(* IEC 61131-3 sources: plc-st-coding-agent/progress/evidence/f14_v14_remaining_20261113/jobs/custom_minimax-m27 (part 9) *)

(* ---- self-medium-04.raw_candidate_01.st ---- *)
FUNCTION_BLOCK FB
VAR_INPUT
    startBtn  : BOOL;
    resetBtn  : BOOL;
    doneSensor: BOOL;
    targetVol : REAL;
    flowVol   : REAL;
END_VAR
VAR_OUTPUT
    valveOpen : BOOL;
    fillsToday: INT;
END_VAR
VAR
    state           : INT;        // 0=IDLE, 1=FILLING, 2=PENDING
    prev_startBtn   : BOOL;
    prev_resetBtn   : BOOL;
    prev_valveOpen  : BOOL;
    pendingConfirm  : BOOL;
    accumulatedVol  : REAL;
    rising_startBtn : BOOL;
    rising_resetBtn : BOOL;
    tmp_doConfirm   : BOOL;
END_VAR

// ENGINEERING_CONTRACT
// States: IDLE(0), FILLING(1), PENDING(2)
// Outputs: valveOpen (BOOL, hold open during FILLING until target reached or reset)
//          fillsToday (INT, hold-until-confirm count, saturation at 32767)
// Confirmed fills increment fillsToday by 1 per bottle, cleared on reset
// ResetBtn rising edge (rising_resetBtn) has absolute priority; clears all state
// StartBtn rising edge (rising_startBtn) in IDLE or PENDING starts new bottle
// Confirmation checks doneSensor at valve-close scan; clears pendingConfirm after
// No hidden timers; all state in VAR; explicit edge detection via prev_* vars

(* CONTRACT_RULES [] *)

rising_startBtn := startBtn AND NOT prev_startBtn;
rising_resetBtn := resetBtn  AND NOT prev_resetBtn;

// PUB001: Reset takes priority - ignore everything else this scan
IF rising_resetBtn THEN
    pendingConfirm := FALSE;
    accumulatedVol := 0.0;
    valveOpen      := FALSE;
    fillsToday     := 0;
    prev_startBtn  := startBtn;
    prev_resetBtn  := resetBtn;
    prev_valveOpen := valveOpen;
    RETURN;
END_IF;

// PUB002: Start new bottle when startBtn rises (idle or waiting confirmation)
IF rising_startBtn AND (state = 0 OR state = 2) THEN
    state           := 1;          // FILLING
    pendingConfirm  := FALSE;      // cancel previous pending if any
    accumulatedVol  := flowVol;    // PUB008: start scan counts flow
    IF accumulatedVol >= targetVol THEN
        valveOpen := FALSE;        // PUB014: immediate达标 close
        tmp_doConfirm := doneSensor;
        IF tmp_doConfirm THEN
            IF fillsToday < 32767 THEN
                fillsToday := fillsToday + 1; // PUB030/PUB031: confirm new bottle
            END_IF;
            pendingConfirm := FALSE;
            state := 0;            // back to idle
        ELSE
            pendingConfirm := TRUE;
            state := 2;            // PENDING
        END_IF;
    ELSE
        valveOpen := TRUE;
    END_IF;
    prev_startBtn  := startBtn;
    prev_resetBtn  := resetBtn;
    prev_valveOpen := valveOpen;
    RETURN;
END_IF;

// PUB003: Accumulate flow during filling, including start scan
IF state = 1 THEN
    accumulatedVol := accumulatedVol + flowVol;
    IF accumulatedVol >= targetVol THEN
        valveOpen := FALSE;
        accumulatedVol := targetVol; // PUB035: cap at target
        pendingConfirm := TRUE;
        tmp_doConfirm := doneSensor;
        IF tmp_doConfirm THEN
            // PUB014/PUB004: 本拍关阀后立即确认
            IF fillsToday < 32767 THEN
                fillsToday := fillsToday + 1;
            END_IF;
            pendingConfirm := FALSE;
            state := 0;
        ELSE
            state := 2; // PUB004: wait for future TRUE
        END_IF;
    END_IF;
END_IF;

// PUB004: In PENDING, confirm on first TRUE of doneSensor (unless reset/start)
IF state = 2 AND doneSensor THEN
    IF fillsToday < 32767 THEN
        fillsToday := fillsToday + 1;
    END_IF;
    pendingConfirm := FALSE;
    state := 0;
END_IF;

// PUB047: New start during PENDING cancels pending before start logic
// Handled above by clearing pendingConfirm on rising_startBtn in PENDING

prev_startBtn  := startBtn;
prev_resetBtn  := resetBtn;
prev_valveOpen := valveOpen;
END_FUNCTION_BLOCK

(* ---- self-medium-04.raw_candidate_03.st ---- *)
FUNCTION_BLOCK FB
VAR_INPUT
    startBtn  : BOOL;
    resetBtn  : BOOL;
    doneSensor: BOOL;
    targetVol : REAL;
    flowVol   : REAL;
END_VAR
VAR_OUTPUT
    valveOpen : BOOL;
    fillsToday: INT;
END_VAR
VAR
    state           : INT;        // 0=IDLE, 1=FILLING, 2=PENDING
    prev_startBtn   : BOOL := FALSE;
    prev_resetBtn   : BOOL := FALSE;
    prev_valveOpen  : BOOL := FALSE;
    pendingConfirm  : BOOL;
    accumulatedVol  : REAL := 0.0;
END_VAR

// ENGINEERING_CONTRACT
// States: IDLE(0), FILLING(1), PENDING(2)
// Outputs: valveOpen (BOOL, hold open during FILLING until target reached or reset)
//          fillsToday (INT, hold-until-confirm count, saturation at 32767)
// Confirmed fills increment fillsToday by 1 per bottle, cleared on reset
// ResetBtn rising edge has absolute priority; clears all state and closes valve
// StartBtn rising edge in IDLE or PENDING starts new bottle, cancels pending
// Confirmation checks doneSensor at valve-close scan; clears pendingConfirm after
// No hidden timers; all state in VAR; explicit edge detection via prev_* vars

(* CONTRACT_RULES [] *)

// PUB001: Reset takes priority - ignore everything else this scan
IF resetBtn AND NOT prev_resetBtn THEN
    pendingConfirm := FALSE;
    accumulatedVol := 0.0;
    valveOpen      := FALSE;
    fillsToday     := 0;
    state          := 0;
    prev_startBtn  := resetBtn;
    prev_resetBtn  := resetBtn;
    prev_valveOpen := valveOpen;
    RETURN;
END_IF;

// PUB002/PUB047: Start new bottle when startBtn rises (idle or waiting confirmation)
IF startBtn AND NOT prev_startBtn AND (state = 0 OR state = 2) THEN
    state          := 1;          // FILLING
    pendingConfirm := FALSE;      // cancel previous pending if any
    accumulatedVol := flowVol;    // PUB008: start scan counts flow
    IF accumulatedVol >= targetVol THEN
        valveOpen := FALSE;        // PUB014: immediate达标 close
        IF doneSensor THEN
            IF fillsToday < 32767 THEN
                fillsToday := fillsToday + 1; // PUB030/PUB031: confirm new bottle
            END_IF;
            pendingConfirm := FALSE;
            state := 0;            // back to idle
        ELSE
            pendingConfirm := TRUE;
            state := 2;            // PENDING
        END_IF;
    ELSE
        valveOpen := TRUE;
    END_IF;
    prev_startBtn  := startBtn;
    prev_resetBtn  := resetBtn;
    prev_valveOpen := valveOpen;
    RETURN;
END_IF;

// PUB003: Accumulate flow during filling, including start scan
IF state = 1 THEN
    accumulatedVol := accumulatedVol + flowVol;
    IF accumulatedVol >= targetVol THEN
        valveOpen := FALSE;
        accumulatedVol := targetVol; // PUB035: cap at target
        pendingConfirm := TRUE;
        IF doneSensor THEN
            // PUB014/PUB004: 本拍关阀后立即确认
            IF fillsToday < 32767 THEN
                fillsToday := fillsToday + 1;
            END_IF;
            pendingConfirm := FALSE;
            state := 0;
        ELSE
            state := 2; // PUB004: wait for future TRUE
        END_IF;
    END_IF;
END_IF;

// PUB004: In PENDING, confirm on first TRUE of doneSensor (unless reset/start)
IF state = 2 AND doneSensor THEN
    IF fillsToday < 32767 THEN
        fillsToday := fillsToday + 1;
    END_IF;
    pendingConfirm := FALSE;
    state := 0;
END_IF;

prev_startBtn  := startBtn;
prev_resetBtn  := resetBtn;
prev_valveOpen := valveOpen;
END_FUNCTION_BLOCK

(* ---- self-medium-05.candidate_01.st ---- *)
(* ENGINEERING_CONTRACT FB_SteamAccumulator
   ┌──────────────┬─────────────────────┬──────────────────────┬───────────────┬─────────────┐
   │ Output       │ Activation          │ Retention            │ Reset/Deact   │ Boundaries  │
   ├──────────────┼─────────────────────┼──────────────────────┼───────────────┼─────────────┤
   │ qualified    │ enable, no fault    │ N/A (combinational)  │ N/A           │ T∈[447,453] │
   │              │                     │                      │               │ P∈[3750,3850]│
   │ dataFault    │ scanSeconds/flow    │ N/A (combinational)  │ N/A           │ dt∈(0,10]   │
   │              │                     │                      │               │ SF∈[0,90]   │
   │              │                     │                      │               │ FF∈[0,6]    │
   │ qualifiedTon │ enable∧no fault∧    │ Hold value on        │ resetBtn↑     │ ≥0, t units │
   │              │ qualified (additive)│ disable/fault/hold   │ clears to 0   │             │
   │ fuelTon      │ enable∧no fault     │ Hold value on        │ resetBtn↑     │ ≥0, t units │
   │              │ (always add)        │ disable/fault/hold   │ clears to 0   │             │
   │ revenue      │ Always updated      │ N/A                  │ N/A           │ ≥0, yuan    │
   │ cost         │ Always updated      │ N/A                  │ N/A           │ ≥0, yuan    │
   │ netProfit    │ Always updated      │ N/A                  │ N/A           │ ±, yuan     │
   └──────────────┴─────────────────────┴──────────────────────┴───────────────┴─────────────┘
   [PUB001] qualified := steamTemp∈[447,453] ∧ steamPressure∈[3750,3850] (closed interval)
   [PUB002] qualifiedTon accumulates when enable∧no fault∧qualified (kg/s×s/1000→t)
   [PUB003] fuelTon always accumulates when enable∧no fault (kg/s×s/1000→t)
   [PUB004] dataFault := scanSeconds≤0 ∨ scanSeconds>10 ∨ steamFlow∉[0,90] ∨ fuelFlow∉[0,6]
   [PUB005] resetBtn↑ → immediate zero, no accumulation in same scan (edge, not level)
   [PUB006] resetBtn↑ takes priority over dataFault; both may report simultaneously
   [PUB007] revenue=qualifiedTon×280, cost=fuelTon×1500, netProfit=revenue-cost (per-scan)
   [PUB008] qualifiedTon/fuelTon/revenue/cost ≥ 0; netProfit may be negative
   [PUB009] No hidden timers; static VAR for state; R_TRIG for edge detection
   [PUB010] same-scan: evaluate final enable/fault before calling accumulation
   [PUB048] Closed-interval qualification; boundary values are QUALIFIED
   [PUB049] ScanSeconds 10.0 is valid; >10.0 is fault
   [PUB050] negative flow values are faults (PUB004 scope)
*)
FUNCTION_BLOCK FB
VAR_INPUT
    enable       : BOOL;
    resetBtn     : BOOL;
    scanSeconds  : LREAL;
    steamFlow    : LREAL;
    fuelFlow     : LREAL;
    steamTemp    : LREAL;
    steamPressure: LREAL;
END_VAR
VAR_OUTPUT
    qualified    : BOOL;
    dataFault    : BOOL;
    qualifiedTon : LREAL;
    fuelTon      : LREAL;
    revenue      : LREAL;
    cost         : LREAL;
    netProfit    : LREAL;
END_VAR
VAR
    resetRtrig   : R_TRIG;
    prevResetBtn : BOOL := FALSE;
    tmpFault     : BOOL;
    tmpEnable    : BOOL;
    tmpAddQ      : LREAL;
    tmpAddF      : LREAL;
END_VAR
VAR_TEMP
    incQualified : LREAL;
    incFuel      : LREAL;
END_VAR
(* ── Scan cycle start ──────────────────────────────────────────────── *)
resetRtrig(CLK := resetBtn);
tmpFault  := (scanSeconds <= 0.0) OR (scanSeconds > 10.0)
              OR (steamFlow < 0.0) OR (steamFlow > 90.0)
              OR (fuelFlow < 0.0)  OR (fuelFlow > 6.0);
tmpEnable := enable AND NOT tmpFault;

qualified := (steamTemp >= 447.0) AND (steamTemp <= 453.0)
             AND (steamPressure >= 3750.0) AND (steamPressure <= 3850.0);

incQualified := 0.0;
incFuel      := 0.0;

(* Accumulation path: only when no reset rising edge this scan *)
IF NOT resetRtrig.Q THEN
    IF tmpEnable THEN
        incFuel := fuelFlow * scanSeconds / 1000.0;
        IF qualified THEN
            incQualified := steamFlow * scanSeconds / 1000.0;
        END_IF;
    END_IF;
    qualifiedTon := qualifiedTon + incQualified;
    fuelTon      := fuelTon + incFuel;
ELSE
    (* Reset rising edge: cleared, no accumulation this scan *)
    qualifiedTon := 0.0;
    fuelTon      := 0.0;
END_IF;

(* Revenue/cost/netProfit: always updated per scan from current accumulators *)
revenue   := qualifiedTon * 280.0;
cost      := fuelTon * 1500.0;
netProfit := revenue - cost;

dataFault := tmpFault;

prevResetBtn := resetBtn;
END_FUNCTION_BLOCK
(* CONTRACT_RULES [] *)

(* ---- self-medium-05.raw_candidate_01.st ---- *)
(* ENGINEERING_CONTRACT FB_SteamAccumulator
   ┌──────────────┬─────────────────────┬──────────────────────┬───────────────┬─────────────┐
   │ Output       │ Activation          │ Retention            │ Reset/Deact   │ Boundaries  │
   ├──────────────┼─────────────────────┼──────────────────────┼───────────────┼─────────────┤
   │ qualified    │ enable, no fault    │ N/A (combinational)  │ N/A           │ T∈[447,453] │
   │              │                     │                      │               │ P∈[3750,3850]│
   │ dataFault    │ scanSeconds/flow    │ N/A (combinational)  │ N/A           │ dt∈(0,10]   │
   │              │                     │                      │               │ SF∈[0,90]   │
   │              │                     │                      │               │ FF∈[0,6]    │
   │ qualifiedTon │ enable∧no fault∧    │ Hold value on        │ resetBtn↑     │ ≥0, t units │
   │              │ qualified (additive)│ disable/fault/hold   │ clears to 0   │             │
   │ fuelTon      │ enable∧no fault     │ Hold value on        │ resetBtn↑     │ ≥0, t units │
   │              │ (always add)        │ disable/fault/hold   │ clears to 0   │             │
   │ revenue      │ Always updated      │ N/A                  │ N/A           │ ≥0, yuan    │
   │ cost         │ Always updated      │ N/A                  │ N/A           │ ≥0, yuan    │
   │ netProfit    │ Always updated      │ N/A                  │ N/A           │ ±, yuan     │
   └──────────────┴─────────────────────┴──────────────────────┴───────────────┴─────────────┘
   [PUB001] qualified := steamTemp∈[447,453] ∧ steamPressure∈[3750,3850] (closed interval)
   [PUB002] qualifiedTon accumulates when enable∧no fault∧qualified (kg/s×s/1000→t)
   [PUB003] fuelTon always accumulates when enable∧no fault (kg/s×s/1000→t)
   [PUB004] dataFault := scanSeconds≤0 ∨ scanSeconds>10 ∨ steamFlow∉[0,90] ∨ fuelFlow∉[0,6]
   [PUB005] resetBtn↑ → immediate zero, no accumulation in same scan (edge, not level)
   [PUB006] resetBtn↑ takes priority over dataFault; both may report simultaneously
   [PUB007] revenue=qualifiedTon×280, cost=fuelTon×1500, netProfit=revenue-cost (per-scan)
   [PUB008] qualifiedTon/fuelTon/revenue/cost ≥ 0; netProfit may be negative
   [PUB009] No hidden timers; static VAR for state; R_TRIG for edge detection
   [PUB010] same-scan: evaluate final enable/fault before calling accumulation
   [PUB048] Closed-interval qualification; boundary values are QUALIFIED
   [PUB049] ScanSeconds 10.0 is valid; >10.0 is fault
   [PUB050] negative flow values are faults (PUB004 scope)
*)
FUNCTION_BLOCK FB
VAR_INPUT
    enable       : BOOL;
    resetBtn     : BOOL;
    scanSeconds  : LREAL;
    steamFlow    : LREAL;
    fuelFlow     : LREAL;
    steamTemp    : LREAL;
    steamPressure: LREAL;
END_VAR
VAR_OUTPUT
    qualified    : BOOL;
    dataFault    : BOOL;
    qualifiedTon : LREAL;
    fuelTon      : LREAL;
    revenue      : LREAL;
    cost         : LREAL;
    netProfit    : LREAL;
END_VAR
VAR
    resetRtrig   : R_TRIG;
    prevResetBtn : BOOL := FALSE;
    tmpFault     : BOOL;
    tmpEnable    : BOOL;
    tmpAddQ      : LREAL;
    tmpAddF      : LREAL;
END_VAR
VAR_TEMP
    incQualified : LREAL;
    incFuel      : LREAL;
END_VAR
(* ── Scan cycle start ──────────────────────────────────────────────── *)
resetRtrig(CLK := resetBtn);
tmpFault  := (scanSeconds <= 0.0) OR (scanSeconds > 10.0)
              OR (steamFlow < 0.0) OR (steamFlow > 90.0)
              OR (fuelFlow < 0.0)  OR (fuelFlow > 6.0);
tmpEnable := enable AND NOT tmpFault;

qualified := (steamTemp >= 447.0) AND (steamTemp <= 453.0)
             AND (steamPressure >= 3750.0) AND (steamPressure <= 3850.0);

incQualified := 0.0;
incFuel      := 0.0;

(* Accumulation path: only when no reset rising edge this scan *)
IF NOT resetRtrig.Q THEN
    IF tmpEnable THEN
        incFuel := fuelFlow * scanSeconds / 1000.0;
        IF qualified THEN
            incQualified := steamFlow * scanSeconds / 1000.0;
        END_IF
    END_IF
    qualifiedTon := qualifiedTon + incQualified;
    fuelTon      := fuelTon + incFuel;
ELSE
    (* Reset rising edge: cleared, no accumulation this scan *)
    qualifiedTon := 0.0;
    fuelTon      := 0.0;
END_IF

(* Revenue/cost/netProfit: always updated per scan from current accumulators *)
revenue   := qualifiedTon * 280.0;
cost      := fuelTon * 1500.0;
netProfit := revenue - cost;

dataFault := tmpFault;

prevResetBtn := resetBtn;
END_FUNCTION_BLOCK
(* CONTRACT_RULES [] *)

(* ---- self-medium-06.candidate_01.st ---- *)
(* ENGINEERING_CONTRACT FB_FuzzyTempControl
   ========================================================================
   Outputs & State Retention:
   --------------------------------------------------------------------
   power:       COMBINATIONAL (bias + correction) clamped to [0,100].
                Zeroed on enable=FALSE, fault=TRUE, or resetBtn rising.
   correction:  COMBINATIONAL weighted-centroid per 9 rules.
                Zeroed same as power; no internal clamping (range ±30).
   fault:       COMBINATIONAL; fault = NOT sensorValid OR scanSeconds
                outside (0,10]. Not latched.
   ePrev:       RETAINED across scans; cleared on rising(resetBtn),
                enable=FALSE, or fault=TRUE.
   tmpHistValid:RETAINED; FALSE after clear, set TRUE after first de.
   tmpResetPrevHigh:RETAINED; set TRUE on rising(resetBtn), cleared
                next scan so held reset allows normal calculation.
   -----------------------------------------------------------------------
   First-scan rule (PUB011/PUB012): when tmpHistValid=FALSE, de=0.
   Subsequent scans use ePrev for differential calculation.
   Reset is edge-triggered only (rising edge clears; held reset allows
   normal fuzzy output per S9).
   ========================================================================
*)
FUNCTION_BLOCK FB
VAR
    ePrev          : REAL := 0.0;
    tmpHistValid   : BOOL := FALSE;
    tmpResetPrevHigh: BOOL := FALSE;
END_VAR
VAR_OUTPUT
    power      : REAL;
    correction : REAL;
    fault      : BOOL;
END_VAR
VAR_INPUT
    enable      : BOOL;
    resetBtn    : BOOL;
    sensorValid : BOOL;
    setpoint    : REAL;
    temperature : REAL;
    scanSeconds : REAL;
    bias        : REAL;
END_VAR

    (* --- Fault determination (PUB004, PUB028) --- *)
    fault := NOT sensorValid OR scanSeconds <= 0.0 OR scanSeconds > 10.0;

    (* --- Reset rising-edge detection (PUB011): edge only, not hold --- *)
    IF resetBtn AND NOT tmpResetPrevHigh THEN
        (* Rising edge of resetBtn this scan: zero outputs, clear history --- *)
        power       := 0.0;
        correction  := 0.0;
        ePrev       := 0.0;
        tmpHistValid := FALSE;
        tmpResetPrevHigh := TRUE;
        RETURN;
    END_IF;

    (* Remember current resetBtn for next-scan edge detection --- *)
    tmpResetPrevHigh := resetBtn;

    (* --- Disabled or faulted: zero outputs, clear history (PUB011) --- *)
    IF NOT enable OR fault THEN
        power       := 0.0;
        correction  := 0.0;
        ePrev       := 0.0;
        tmpHistValid := FALSE;
        RETURN;
    END_IF;

    (* ==================================================================
       Normal fuzzy calculation
       ================================================================== *)
    VAR
        e          : REAL;
        de         : REAL;
        x          : REAL;
        y          : REAL;
        muN_x      : REAL;
        muZ_x      : REAL;
        muP_x      : REAL;
        muN_y      : REAL;
        muZ_y      : REAL;
        muP_y      : REAL;
        w           : ARRAY[1..3, 1..3] OF REAL;
        sumW        : REAL;
        sumWc       : REAL;
        row         : INT;
        col         : INT;
        tmpFirstScan: BOOL;
    END_VAR

    (* PUB001: error definition --- *)
    e := setpoint - temperature;

    (* PUB012: first-scan detection --- *)
    tmpFirstScan := NOT tmpHistValid;

    (* PUB011: de = 0 on first scan or after history clear --- *)
    IF tmpFirstScan THEN
        de := 0.0;
    ELSE
        de := (e - ePrev) / scanSeconds;
    END_IF;

    (* PUB003 / PUB005: normalize to [-1,1] --- *)
    x := LIMIT(-1.0, e / 10.0, 1.0);
    y := LIMIT(-1.0, de / 2.0, 1.0);

    (* PUB006: membership functions --- *)
    muN_x := MAX(-x, 0.0);
    muZ_x := MAX(1.0 - ABS(x), 0.0);
    muP_x := MAX( x, 0.0);

    muN_y := MAX(-y, 0.0);
    muZ_y := MAX(1.0 - ABS(y), 0.0);
    muP_y := MAX( y, 0.0);

    (* Rule weights: row = x (N/Z/P), col = y (N/Z/P) --- *)
    w[1,1] := muN_x * muN_y;   (* N,N *)
    w[1,2] := muN_x * muZ_y;   (* N,Z *)
    w[1,3] := muN_x * muP_y;   (* N,P *)
    w[2,1] := muZ_x * muN_y;   (* Z,N *)
    w[2,2] := muZ_x * muZ_y;   (* Z,Z *)
    w[2,3] := muZ_x * muP_y;   (* Z,P *)
    w[3,1] := muP_x * muN_y;   (* P,N *)
    w[3,2] := muP_x * muZ_y;   (* P,Z *)
    w[3,3] := muP_x * muP_y;   (* P,P *)

    (* Weighted centroid (PUB007): sum(w*c)/sum(w) --- *)
    sumW  := 0.0;
    sumWc := 0.0;
    FOR row := 1 TO 3 DO
        FOR col := 1 TO 3 DO
            sumW  := sumW  + w[row, col];
            sumWc := sumWc + w[row, col] * SEL(INT_TO_INT(row - 1), SEL(INT_TO_INT(col - 1),
                                 -30.0,   (* row=1 (N) *)
                                 -10.0,   (* row=2 (Z) *)
                                  10.0),  (* row=3 (P) *)
                                 SEL(INT_TO_INT(col - 1),
                                 -20.0,   (* col=1 (N) *)
                                   0.0,   (* col=2 (Z) *)
                                  20.0)); (* col=3 (P) *)
        END_FOR;
    END_FOR;

    (* PUB007: Σw=0 → correction=0 --- *)
    IF sumW > 0.0 THEN
        correction := sumWc / sumW;
    ELSE
        correction := 0.0;
    END_IF;

    (* PUB008: power = clamp(bias + correction, 0, 100) --- *)
    power := LIMIT(0.0, bias + correction, 100.0);

    (* Update history for next scan --- *)
    ePrev       := e;
    tmpHistValid := TRUE;
END_FUNCTION_BLOCK

(* ---- self-medium-06.candidate_03.st ---- *)
(* ENGINEERING_CONTRACT FB_FuzzyTempControl
   ========================================================================
   Outputs & State Retention:
   --------------------------------------------------------------------
   power:       COMBINATIONAL (bias + correction) clamped to [0,100].
                Zeroed on enable=FALSE, fault=TRUE, or resetBtn rising.
   correction:  COMBINATIONAL weighted-centroid per 9 rules.
                Zeroed same as power; no internal clamping (range ±30).
   fault:       COMBINATIONAL; fault = NOT sensorValid OR scanSeconds
                outside (0,10]. Not latched.
   ePrev:       RETAINED across scans; cleared on rising(resetBtn),
                enable=FALSE, or fault=TRUE.
   tmpHistValid:RETAINED; FALSE after clear, set TRUE after first de.
   tmpResetPrevHigh:RETAINED; set TRUE on rising(resetBtn), cleared
                next scan so held reset allows normal calculation.
   -----------------------------------------------------------------------
   First-scan rule (PUB011/PUB012): when tmpHistValid=FALSE, de=0.
   Subsequent scans use ePrev for differential calculation.
   Reset is edge-triggered only (rising edge clears; held reset allows
   normal fuzzy output per S9).
   ========================================================================
*)
FUNCTION_BLOCK FB
VAR
    ePrev          : REAL := 0.0;
    tmpHistValid   : BOOL := FALSE;
    tmpResetPrevHigh: BOOL := FALSE;
END_VAR
VAR_OUTPUT
    power      : REAL;
    correction : REAL;
    fault      : BOOL;
END_VAR
VAR_INPUT
    enable      : BOOL;
    resetBtn    : BOOL;
    sensorValid : BOOL;
    setpoint    : REAL;
    temperature : REAL;
    scanSeconds : REAL;
    bias        : REAL;
END_VAR

    (* --- Fault determination (PUB004, PUB028) --- *)
    fault := NOT sensorValid OR scanSeconds <= 0.0 OR scanSeconds > 10.0;

    (* --- Reset rising-edge detection (PUB011): edge only, not hold --- *)
    IF resetBtn AND NOT tmpResetPrevHigh THEN
        (* Rising edge of resetBtn this scan: zero outputs, clear history --- *)
        power       := 0.0;
        correction  := 0.0;
        ePrev       := 0.0;
        tmpHistValid := FALSE;
        tmpResetPrevHigh := TRUE;
        RETURN;
    END_IF;

    (* Remember current resetBtn for next-scan edge detection --- *)
    tmpResetPrevHigh := resetBtn;

    (* --- Disabled or faulted: zero outputs, clear history (PUB011) --- *)
    IF NOT enable OR fault THEN
        power       := 0.0;
        correction  := 0.0;
        ePrev       := 0.0;
        tmpHistValid := FALSE;
        RETURN;
    END_IF;

    (* ==================================================================
       Normal fuzzy calculation
       ================================================================== *)
    (* local computation variables *)
    e           : REAL;
    de          : REAL;
    x           : REAL;
    y           : REAL;
    muN_x       : REAL;
    muZ_x       : REAL;
    muP_x       : REAL;
    muN_y       : REAL;
    muZ_y       : REAL;
    muP_y       : REAL;
    w           : ARRAY[1..3, 1..3] OF REAL;
    sumW        : REAL;
    sumWc       : REAL;
    row         : INT;
    col         : INT;
    tmpFirstScan: BOOL;
END_VAR

    (* PUB001: error definition --- *)
    e := setpoint - temperature;

    (* PUB012: first-scan detection --- *)
    tmpFirstScan := NOT tmpHistValid;

    (* PUB011: de = 0 on first scan or after history clear --- *)
    IF tmpFirstScan THEN
        de := 0.0;
    ELSE
        de := (e - ePrev) / scanSeconds;
    END_IF;

    (* PUB003 / PUB005: normalize to [-1,1] --- *)
    x := LIMIT(-1.0, e / 10.0, 1.0);
    y := LIMIT(-1.0, de / 2.0, 1.0);

    (* PUB006: membership functions --- *)
    muN_x := MAX(-x, 0.0);
    muZ_x := MAX(1.0 - ABS(x), 0.0);
    muP_x := MAX( x, 0.0);

    muN_y := MAX(-y, 0.0);
    muZ_y := MAX(1.0 - ABS(y), 0.0);
    muP_y := MAX( y, 0.0);

    (* Rule weights: row = x (N/Z/P), col = y (N/Z/P) --- *)
    w[1,1] := muN_x * muN_y;   (* N,N *)
    w[1,2] := muN_x * muZ_y;   (* N,Z *)
    w[1,3] := muN_x * muP_y;   (* N,P *)
    w[2,1] := muZ_x * muN_y;   (* Z,N *)
    w[2,2] := muZ_x * muZ_y;   (* Z,Z *)
    w[2,3] := muZ_x * muP_y;   (* Z,P *)
    w[3,1] := muP_x * muN_y;   (* P,N *)
    w[3,2] := muP_x * muZ_y;   (* P,Z *)
    w[3,3] := muP_x * muP_y;   (* P,P *)

    (* Weighted centroid (PUB007): sum(w*c)/sum(w) --- *)
    sumW  := 0.0;
    sumWc := 0.0;
    FOR row := 1 TO 3 DO
        FOR col := 1 TO 3 DO
            sumW  := sumW  + w[row, col];
            sumWc := sumWc + w[row, col] * SEL(INT_TO_INT(row - 1), SEL(INT_TO_INT(col - 1),
                                 -30.0,   (* row=1 (N) *)
                                 -10.0,   (* row=2 (Z) *)
                                  10.0),  (* row=3 (P) *)
                                 SEL(INT_TO_INT(col - 1),
                                 -20.0,   (* col=1 (N) *)
                                   0.0,   (* col=2 (Z) *)
                                  20.0)); (* col=3 (P) *)
        END_FOR;
    END_FOR;

    (* PUB007: Σw=0 → correction=0 --- *)
    IF sumW > 0.0 THEN
        correction := sumWc / sumW;
    ELSE
        correction := 0.0;
    END_IF;

    (* PUB008: power = clamp(bias + correction, 0, 100) --- *)
    power := LIMIT(0.0, bias + correction, 100.0);

    (* Update history for next scan --- *)
    ePrev       := e;
    tmpHistValid := TRUE;
END_FUNCTION_BLOCK

(* ---- self-medium-06.candidate_04.st ---- *)
(* ENGINEERING_CONTRACT FB_FuzzyTempControl
   ========================================================================
   Outputs & State Retention:
   --------------------------------------------------------------------
   power:       COMBINATIONAL (bias + correction) clamped to [0,100].
                Zeroed on enable=FALSE, fault=TRUE, or resetBtn rising.
   correction:  COMBINATIONAL weighted-centroid per 9 rules.
                Zeroed same as power; no internal clamping (range ±30).
   fault:       COMBINATIONAL; fault = NOT sensorValid OR scanSeconds
                outside (0,10]. Not latched.
   ePrev:       RETAINED across scans; cleared on rising(resetBtn),
                enable=FALSE, or fault=TRUE.
   tmpHistValid:RETAINED; FALSE after clear, set TRUE after first de.
   tmpResetPrevHigh:RETAINED; set TRUE on rising(resetBtn), cleared
                next scan so held reset allows normal calculation.
   -----------------------------------------------------------------------
   First-scan rule (PUB011/PUB012): when tmpHistValid=FALSE, de=0.
   Subsequent scans use ePrev for differential calculation.
   Reset is edge-triggered only (rising edge clears; held reset allows
   normal fuzzy output per S9).
   ========================================================================
*)
FUNCTION_BLOCK FB
VAR
    ePrev           : REAL := 0.0;
    tmpHistValid    : BOOL := FALSE;
    tmpResetPrevHigh: BOOL := FALSE;
    e               : REAL;
    de              : REAL;
    x               : REAL;
    y               : REAL;
    muN_x           : REAL;
    muZ_x           : REAL;
    muP_x           : REAL;
    muN_y           : REAL;
    muZ_y           : REAL;
    muP_y           : REAL;
    w               : ARRAY[1..3, 1..3] OF REAL;
    sumW            : REAL;
    sumWc           : REAL;
    row             : INT;
    col             : INT;
    tmpFirstScan    : BOOL;
END_VAR
VAR_OUTPUT
    power      : REAL;
    correction : REAL;
    fault      : BOOL;
END_VAR
VAR_INPUT
    enable      : BOOL;
    resetBtn    : BOOL;
    sensorValid : BOOL;
    setpoint    : REAL;
    temperature : REAL;
    scanSeconds : REAL;
    bias        : REAL;
END_VAR

    (* --- Fault determination (PUB004, PUB028) --- *)
    fault := NOT sensorValid OR scanSeconds <= 0.0 OR scanSeconds > 10.0;

    (* --- Reset rising-edge detection (PUB011): edge only, not hold --- *)
    IF resetBtn AND NOT tmpResetPrevHigh THEN
        (* Rising edge of resetBtn this scan: zero outputs, clear history --- *)
        power        := 0.0;
        correction   := 0.0;
        ePrev        := 0.0;
        tmpHistValid := FALSE;
        tmpResetPrevHigh := TRUE;
        RETURN;
    END_IF;

    (* Remember current resetBtn for next-scan edge detection --- *)
    tmpResetPrevHigh := resetBtn;

    (* --- Disabled or faulted: zero outputs, clear history (PUB011) --- *)
    IF NOT enable OR fault THEN
        power        := 0.0;
        correction   := 0.0;
        ePrev        := 0.0;
        tmpHistValid := FALSE;
        RETURN;
    END_IF;

    (* ==================================================================
       Normal fuzzy calculation
       ================================================================== *)

    (* PUB001: error definition --- *)
    e := setpoint - temperature;

    (* PUB012: first-scan detection --- *)
    tmpFirstScan := NOT tmpHistValid;

    (* PUB011: de = 0 on first scan or after history clear --- *)
    IF tmpFirstScan THEN
        de := 0.0;
    ELSE
        de := (e - ePrev) / scanSeconds;
    END_IF;

    (* PUB003 / PUB005: normalize to [-1,1] --- *)
    x := LIMIT(-1.0, e / 10.0, 1.0);
    y := LIMIT(-1.0, de / 2.0, 1.0);

    (* PUB006: membership functions --- *)
    muN_x := MAX(-x, 0.0);
    muZ_x := MAX(1.0 - ABS(x), 0.0);
    muP_x := MAX( x, 0.0);

    muN_y := MAX(-y, 0.0);
    muZ_y := MAX(1.0 - ABS(y), 0.0);
    muP_y := MAX( y, 0.0);

    (* Rule weights: row = x (N/Z/P), col = y (N/Z/P) --- *)
    w[1,1] := muN_x * muN_y;   (* N,N *)
    w[1,2] := muN_x * muZ_y;   (* N,Z *)
    w[1,3] := muN_x * muP_y;   (* N,P *)
    w[2,1] := muZ_x * muN_y;   (* Z,N *)
    w[2,2] := muZ_x * muZ_y;   (* Z,Z *)
    w[2,3] := muZ_x * muP_y;   (* Z,P *)
    w[3,1] := muP_x * muN_y;   (* P,N *)
    w[3,2] := muP_x * muZ_y;   (* P,Z *)
    w[3,3] := muP_x * muP_y;   (* P,P *)

    (* Weighted centroid (PUB007): sum(w*c)/sum(w) --- *)
    sumW  := 0.0;
    sumWc := 0.0;
    FOR row := 1 TO 3 DO
        FOR col := 1 TO 3 DO
            sumW  := sumW  + w[row, col];
            sumWc := sumWc + w[row, col] * SEL(INT_TO_INT(row - 1), SEL(INT_TO_INT(col - 1),
                                 -30.0,   (* row=1 (N) *)
                                 -10.0,   (* row=2 (Z) *)
                                  10.0),  (* row=3 (P) *)
                                 SEL(INT_TO_INT(col - 1),
                                 -20.0,   (* col=1 (N) *)
                                   0.0,   (* col=2 (Z) *)
                                  20.0)); (* col=3 (P) *)
        END_FOR;
    END_FOR;

    (* PUB007: Σw=0 → correction=0 --- *)
    IF sumW > 0.0 THEN
        correction := sumWc / sumW;
    ELSE
        correction := 0.0;
    END_IF;

    (* PUB008: power = clamp(bias + correction, 0, 100) --- *)
    power := LIMIT(0.0, bias + correction, 100.0);

    (* Update history for next scan --- *)
    ePrev        := e;
    tmpHistValid := TRUE;
END_FUNCTION_BLOCK

(* ---- self-medium-06.patch_base_02.st ---- *)
(* ENGINEERING_CONTRACT FB_FuzzyTempControl
   ========================================================================
   Outputs & State Retention:
   --------------------------------------------------------------------
   power:       COMBINATIONAL (bias + correction) clamped to [0,100].
                Zeroed on enable=FALSE, fault=TRUE, or resetBtn rising.
   correction:  COMBINATIONAL weighted-centroid per 9 rules.
                Zeroed same as power; no internal clamping (range ±30).
   fault:       COMBINATIONAL; fault = NOT sensorValid OR scanSeconds
                outside (0,10]. Not latched.
   ePrev:       RETAINED across scans; cleared on rising(resetBtn),
                enable=FALSE, or fault=TRUE.
   tmpHistValid:RETAINED; FALSE after clear, set TRUE after first de.
   tmpResetPrevHigh:RETAINED; set TRUE on rising(resetBtn), cleared
                next scan so held reset allows normal calculation.
   -----------------------------------------------------------------------
   First-scan rule (PUB011/PUB012): when tmpHistValid=FALSE, de=0.
   Subsequent scans use ePrev for differential calculation.
   Reset is edge-triggered only (rising edge clears; held reset allows
   normal fuzzy output per S9).
   ========================================================================
*)
FUNCTION_BLOCK FB
VAR
    ePrev          : REAL := 0.0;
    tmpHistValid   : BOOL := FALSE;
    tmpResetPrevHigh: BOOL := FALSE;
END_VAR
VAR_OUTPUT
    power      : REAL;
    correction : REAL;
    fault      : BOOL;
END_VAR
VAR_INPUT
    enable      : BOOL;
    resetBtn    : BOOL;
    sensorValid : BOOL;
    setpoint    : REAL;
    temperature : REAL;
    scanSeconds : REAL;
    bias        : REAL;
END_VAR

    (* --- Fault determination (PUB004, PUB028) --- *)
    fault := NOT sensorValid OR scanSeconds <= 0.0 OR scanSeconds > 10.0;

    (* --- Reset rising-edge detection (PUB011): edge only, not hold --- *)
    IF resetBtn AND NOT tmpResetPrevHigh THEN
        (* Rising edge of resetBtn this scan: zero outputs, clear history --- *)
        power       := 0.0;
        correction  := 0.0;
        ePrev       := 0.0;
        tmpHistValid := FALSE;
        tmpResetPrevHigh := TRUE;
        RETURN;
    END_IF;

    (* Remember current resetBtn for next-scan edge detection --- *)
    tmpResetPrevHigh := resetBtn;

    (* --- Disabled or faulted: zero outputs, clear history (PUB011) --- *)
    IF NOT enable OR fault THEN
        power       := 0.0;
        correction  := 0.0;
        ePrev       := 0.0;
        tmpHistValid := FALSE;
        RETURN;
    END_IF;

    (* ==================================================================
       Normal fuzzy calculation
       ================================================================== *)
    VAR
        e          : REAL;
        de         : REAL;
        x          : REAL;
        y          : REAL;
        muN_x      : REAL;
        muZ_x      : REAL;
        muP_x      : REAL;
        muN_y      : REAL;
        muZ_y      : REAL;
        muP_y      : REAL;
        w           : ARRAY[1..3, 1..3] OF REAL;
        sumW        : REAL;
        sumWc       : REAL;
        row         : INT;
        col         : INT;
        tmpFirstScan: BOOL;
    END_VAR

    (* PUB001: error definition --- *)
    e := setpoint - temperature;

    (* PUB012: first-scan detection --- *)
    tmpFirstScan := NOT tmpHistValid;

    (* PUB011: de = 0 on first scan or after history clear --- *)
    IF tmpFirstScan THEN
        de := 0.0;
    ELSE
        de := (e - ePrev) / scanSeconds;
    END_IF;

    (* PUB003 / PUB005: normalize to [-1,1] --- *)
    x := LIMIT(-1.0, e / 10.0, 1.0);
    y := LIMIT(-1.0, de / 2.0, 1.0);

    (* PUB006: membership functions --- *)
    muN_x := MAX(-x, 0.0);
    muZ_x := MAX(1.0 - ABS(x), 0.0);
    muP_x := MAX( x, 0.0);

    muN_y := MAX(-y, 0.0);
    muZ_y := MAX(1.0 - ABS(y), 0.0);
    muP_y := MAX( y, 0.0);

    (* Rule weights: row = x (N/Z/P), col = y (N/Z/P) --- *)
    w[1,1] := muN_x * muN_y;   (* N,N *)
    w[1,2] := muN_x * muZ_y;   (* N,Z *)
    w[1,3] := muN_x * muP_y;   (* N,P *)
    w[2,1] := muZ_x * muN_y;   (* Z,N *)
    w[2,2] := muZ_x * muZ_y;   (* Z,Z *)
    w[2,3] := muZ_x * muP_y;   (* Z,P *)
    w[3,1] := muP_x * muN_y;   (* P,N *)
    w[3,2] := muP_x * muZ_y;   (* P,Z *)
    w[3,3] := muP_x * muP_y;   (* P,P *)

    (* Weighted centroid (PUB007): sum(w*c)/sum(w) --- *)
    sumW  := 0.0;
    sumWc := 0.0;
    FOR row := 1 TO 3 DO
        FOR col := 1 TO 3 DO
            sumW  := sumW  + w[row, col];
            sumWc := sumWc + w[row, col] * SEL(INT_TO_INT(row - 1), SEL(INT_TO_INT(col - 1),
                                 -30.0,   (* row=1 (N) *)
                                 -10.0,   (* row=2 (Z) *)
                                  10.0),  (* row=3 (P) *)
                                 SEL(INT_TO_INT(col - 1),
                                 -20.0,   (* col=1 (N) *)
                                   0.0,   (* col=2 (Z) *)
                                  20.0)); (* col=3 (P) *)
        END_FOR;
    END_FOR;

    (* PUB007: Σw=0 → correction=0 --- *)
    IF sumW > 0.0 THEN
        correction := sumWc / sumW;
    ELSE
        correction := 0.0;
    END_IF;

    (* PUB008: power = clamp(bias + correction, 0, 100) --- *)
    power := LIMIT(0.0, bias + correction, 100.0);

    (* Update history for next scan --- *)
    ePrev       := e;
    tmpHistValid := TRUE;
END_FUNCTION_BLOCK

(* ---- self-medium-06.patch_base_03.st ---- *)
(* ENGINEERING_CONTRACT FB_FuzzyTempControl
   ========================================================================
   Outputs & State Retention:
   --------------------------------------------------------------------
   power:       COMBINATIONAL (bias + correction) clamped to [0,100].
                Zeroed on enable=FALSE, fault=TRUE, or resetBtn rising.
   correction:  COMBINATIONAL weighted-centroid per 9 rules.
                Zeroed same as power; no internal clamping (range ±30).
   fault:       COMBINATIONAL; fault = NOT sensorValid OR scanSeconds
                outside (0,10]. Not latched.
   ePrev:       RETAINED across scans; cleared on rising(resetBtn),
                enable=FALSE, or fault=TRUE.
   tmpHistValid:RETAINED; FALSE after clear, set TRUE after first de.
   tmpResetPrevHigh:RETAINED; set TRUE on rising(resetBtn), cleared
                next scan so held reset allows normal calculation.
   -----------------------------------------------------------------------
   First-scan rule (PUB011/PUB012): when tmpHistValid=FALSE, de=0.
   Subsequent scans use ePrev for differential calculation.
   Reset is edge-triggered only (rising edge clears; held reset allows
   normal fuzzy output per S9).
   ========================================================================
*)
FUNCTION_BLOCK FB
VAR
    ePrev          : REAL := 0.0;
    tmpHistValid   : BOOL := FALSE;
    tmpResetPrevHigh: BOOL := FALSE;
END_VAR
VAR_OUTPUT
    power      : REAL;
    correction : REAL;
    fault      : BOOL;
END_VAR
VAR_INPUT
    enable      : BOOL;
    resetBtn    : BOOL;
    sensorValid : BOOL;
    setpoint    : REAL;
    temperature : REAL;
    scanSeconds : REAL;
    bias        : REAL;
END_VAR

    (* --- Fault determination (PUB004, PUB028) --- *)
    fault := NOT sensorValid OR scanSeconds <= 0.0 OR scanSeconds > 10.0;

    (* --- Reset rising-edge detection (PUB011): edge only, not hold --- *)
    IF resetBtn AND NOT tmpResetPrevHigh THEN
        (* Rising edge of resetBtn this scan: zero outputs, clear history --- *)
        power       := 0.0;
        correction  := 0.0;
        ePrev       := 0.0;
        tmpHistValid := FALSE;
        tmpResetPrevHigh := TRUE;
        RETURN;
    END_IF;

    (* Remember current resetBtn for next-scan edge detection --- *)
    tmpResetPrevHigh := resetBtn;

    (* --- Disabled or faulted: zero outputs, clear history (PUB011) --- *)
    IF NOT enable OR fault THEN
        power       := 0.0;
        correction  := 0.0;
        ePrev       := 0.0;
        tmpHistValid := FALSE;
        RETURN;
    END_IF;

    (* ==================================================================
       Normal fuzzy calculation
       ================================================================== *)
    VAR
        e          : REAL;
        de         : REAL;
        x          : REAL;
        y          : REAL;
        muN_x      : REAL;
        muZ_x      : REAL;
        muP_x      : REAL;
        muN_y      : REAL;
        muZ_y      : REAL;
        muP_y      : REAL;
        w           : ARRAY[1..3, 1..3] OF REAL;
        sumW        : REAL;
        sumWc       : REAL;
        row         : INT;
        col         : INT;
        tmpFirstScan: BOOL;
    END_VAR

    (* PUB001: error definition --- *)
    e := setpoint - temperature;

    (* PUB012: first-scan detection --- *)
    tmpFirstScan := NOT tmpHistValid;

    (* PUB011: de = 0 on first scan or after history clear --- *)
    IF tmpFirstScan THEN
        de := 0.0;
    ELSE
        de := (e - ePrev) / scanSeconds;
    END_IF;

    (* PUB003 / PUB005: normalize to [-1,1] --- *)
    x := LIMIT(-1.0, e / 10.0, 1.0);
    y := LIMIT(-1.0, de / 2.0, 1.0);

    (* PUB006: membership functions --- *)
    muN_x := MAX(-x, 0.0);
    muZ_x := MAX(1.0 - ABS(x), 0.0);
    muP_x := MAX( x, 0.0);

    muN_y := MAX(-y, 0.0);
    muZ_y := MAX(1.0 - ABS(y), 0.0);
    muP_y := MAX( y, 0.0);

    (* Rule weights: row = x (N/Z/P), col = y (N/Z/P) --- *)
    w[1,1] := muN_x * muN_y;   (* N,N *)
    w[1,2] := muN_x * muZ_y;   (* N,Z *)
    w[1,3] := muN_x * muP_y;   (* N,P *)
    w[2,1] := muZ_x * muN_y;   (* Z,N *)
    w[2,2] := muZ_x * muZ_y;   (* Z,Z *)
    w[2,3] := muZ_x * muP_y;   (* Z,P *)
    w[3,1] := muP_x * muN_y;   (* P,N *)
    w[3,2] := muP_x * muZ_y;   (* P,Z *)
    w[3,3] := muP_x * muP_y;   (* P,P *)

    (* Weighted centroid (PUB007): sum(w*c)/sum(w) --- *)
    sumW  := 0.0;
    sumWc := 0.0;
    FOR row := 1 TO 3 DO
        FOR col := 1 TO 3 DO
            sumW  := sumW  + w[row, col];
            sumWc := sumWc + w[row, col] * SEL(INT_TO_INT(row - 1), SEL(INT_TO_INT(col - 1),
                                 -30.0,   (* row=1 (N) *)
                                 -10.0,   (* row=2 (Z) *)
                                  10.0),  (* row=3 (P) *)
                                 SEL(INT_TO_INT(col - 1),
                                 -20.0,   (* col=1 (N) *)
                                   0.0,   (* col=2 (Z) *)
                                  20.0)); (* col=3 (P) *)
        END_FOR;
    END_FOR;

    (* PUB007: Σw=0 → correction=0 --- *)
    IF sumW > 0.0 THEN
        correction := sumWc / sumW;
    ELSE
        correction := 0.0;
    END_IF;

    (* PUB008: power = clamp(bias + correction, 0, 100) --- *)
    power := LIMIT(0.0, bias + correction, 100.0);

    (* Update history for next scan --- *)
    ePrev       := e;
    tmpHistValid := TRUE;
END_FUNCTION_BLOCK

(* ---- self-medium-06.patch_base_04.st ---- *)
(* ENGINEERING_CONTRACT FB_FuzzyTempControl
   ========================================================================
   Outputs & State Retention:
   --------------------------------------------------------------------
   power:       COMBINATIONAL (bias + correction) clamped to [0,100].
                Zeroed on enable=FALSE, fault=TRUE, or resetBtn rising.
   correction:  COMBINATIONAL weighted-centroid per 9 rules.
                Zeroed same as power; no internal clamping (range ±30).
   fault:       COMBINATIONAL; fault = NOT sensorValid OR scanSeconds
                outside (0,10]. Not latched.
   ePrev:       RETAINED across scans; cleared on rising(resetBtn),
                enable=FALSE, or fault=TRUE.
   tmpHistValid:RETAINED; FALSE after clear, set TRUE after first de.
   tmpResetPrevHigh:RETAINED; set TRUE on rising(resetBtn), cleared
                next scan so held reset allows normal calculation.
   -----------------------------------------------------------------------
   First-scan rule (PUB011/PUB012): when tmpHistValid=FALSE, de=0.
   Subsequent scans use ePrev for differential calculation.
   Reset is edge-triggered only (rising edge clears; held reset allows
   normal fuzzy output per S9).
   ========================================================================
*)
FUNCTION_BLOCK FB
VAR
    ePrev          : REAL := 0.0;
    tmpHistValid   : BOOL := FALSE;
    tmpResetPrevHigh: BOOL := FALSE;
END_VAR
VAR_OUTPUT
    power      : REAL;
    correction : REAL;
    fault      : BOOL;
END_VAR
VAR_INPUT
    enable      : BOOL;
    resetBtn    : BOOL;
    sensorValid : BOOL;
    setpoint    : REAL;
    temperature : REAL;
    scanSeconds : REAL;
    bias        : REAL;
END_VAR

    (* --- Fault determination (PUB004, PUB028) --- *)
    fault := NOT sensorValid OR scanSeconds <= 0.0 OR scanSeconds > 10.0;

    (* --- Reset rising-edge detection (PUB011): edge only, not hold --- *)
    IF resetBtn AND NOT tmpResetPrevHigh THEN
        (* Rising edge of resetBtn this scan: zero outputs, clear history --- *)
        power       := 0.0;
        correction  := 0.0;
        ePrev       := 0.0;
        tmpHistValid := FALSE;
        tmpResetPrevHigh := TRUE;
        RETURN;
    END_IF;

    (* Remember current resetBtn for next-scan edge detection --- *)
    tmpResetPrevHigh := resetBtn;

    (* --- Disabled or faulted: zero outputs, clear history (PUB011) --- *)
    IF NOT enable OR fault THEN
        power       := 0.0;
        correction  := 0.0;
        ePrev       := 0.0;
        tmpHistValid := FALSE;
        RETURN;
    END_IF;

    (* ==================================================================
       Normal fuzzy calculation
       ================================================================== *)
    VAR
        e          : REAL;
        de         : REAL;
        x          : REAL;
        y          : REAL;
        muN_x      : REAL;
        muZ_x      : REAL;
        muP_x      : REAL;
        muN_y      : REAL;
        muZ_y      : REAL;
        muP_y      : REAL;
        w           : ARRAY[1..3, 1..3] OF REAL;
        sumW        : REAL;
        sumWc       : REAL;
        row         : INT;
        col         : INT;
        tmpFirstScan: BOOL;
    END_VAR

    (* PUB001: error definition --- *)
    e := setpoint - temperature;

    (* PUB012: first-scan detection --- *)
    tmpFirstScan := NOT tmpHistValid;

    (* PUB011: de = 0 on first scan or after history clear --- *)
    IF tmpFirstScan THEN
        de := 0.0;
    ELSE
        de := (e - ePrev) / scanSeconds;
    END_IF;

    (* PUB003 / PUB005: normalize to [-1,1] --- *)
    x := LIMIT(-1.0, e / 10.0, 1.0);
    y := LIMIT(-1.0, de / 2.0, 1.0);

    (* PUB006: membership functions --- *)
    muN_x := MAX(-x, 0.0);
    muZ_x := MAX(1.0 - ABS(x), 0.0);
    muP_x := MAX( x, 0.0);

    muN_y := MAX(-y, 0.0);
    muZ_y := MAX(1.0 - ABS(y), 0.0);
    muP_y := MAX( y, 0.0);

    (* Rule weights: row = x (N/Z/P), col = y (N/Z/P) --- *)
    w[1,1] := muN_x * muN_y;   (* N,N *)
    w[1,2] := muN_x * muZ_y;   (* N,Z *)
    w[1,3] := muN_x * muP_y;   (* N,P *)
    w[2,1] := muZ_x * muN_y;   (* Z,N *)
    w[2,2] := muZ_x * muZ_y;   (* Z,Z *)
    w[2,3] := muZ_x * muP_y;   (* Z,P *)
    w[3,1] := muP_x * muN_y;   (* P,N *)
    w[3,2] := muP_x * muZ_y;   (* P,Z *)
    w[3,3] := muP_x * muP_y;   (* P,P *)

    (* Weighted centroid (PUB007): sum(w*c)/sum(w) --- *)
    sumW  := 0.0;
    sumWc := 0.0;
    FOR row := 1 TO 3 DO
        FOR col := 1 TO 3 DO
            sumW  := sumW  + w[row, col];
            sumWc := sumWc + w[row, col] * SEL(INT_TO_INT(row - 1), SEL(INT_TO_INT(col - 1),
                                 -30.0,   (* row=1 (N) *)
                                 -10.0,   (* row=2 (Z) *)
                                  10.0),  (* row=3 (P) *)
                                 SEL(INT_TO_INT(col - 1),
                                 -20.0,   (* col=1 (N) *)
                                   0.0,   (* col=2 (Z) *)
                                  20.0)); (* col=3 (P) *)
        END_FOR;
    END_FOR;

    (* PUB007: Σw=0 → correction=0 --- *)
    IF sumW > 0.0 THEN
        correction := sumWc / sumW;
    ELSE
        correction := 0.0;
    END_IF;

    (* PUB008: power = clamp(bias + correction, 0, 100) --- *)
    power := LIMIT(0.0, bias + correction, 100.0);

    (* Update history for next scan --- *)
    ePrev       := e;
    tmpHistValid := TRUE;
END_FUNCTION_BLOCK

(* ---- self-medium-06.raw_candidate_01.st ---- *)
(* ENGINEERING_CONTRACT FB_FuzzyTempControl
   ========================================================================
   Outputs & State Retention:
   --------------------------------------------------------------------
   power:       COMBINATIONAL (bias + correction) clamped to [0,100].
                Zeroed on enable=FALSE, fault=TRUE, or resetBtn rising.
   correction:  COMBINATIONAL weighted-centroid per 9 rules.
                Zeroed same as power; no internal clamping (range ±30).
   fault:       COMBINATIONAL; fault = NOT sensorValid OR scanSeconds
                outside (0,10]. Not latched.
   ePrev:       RETAINED across scans; cleared on rising(resetBtn),
                enable=FALSE, or fault=TRUE.
   tmpHistValid:RETAINED; FALSE after clear, set TRUE after first de.
   tmpResetPrevHigh:RETAINED; set TRUE on rising(resetBtn), cleared
                next scan so held reset allows normal calculation.
   -----------------------------------------------------------------------
   First-scan rule (PUB011/PUB012): when tmpHistValid=FALSE, de=0.
   Subsequent scans use ePrev for differential calculation.
   Reset is edge-triggered only (rising edge clears; held reset allows
   normal fuzzy output per S9).
   ========================================================================
*)
FUNCTION_BLOCK FB
VAR
    ePrev          : REAL := 0.0;
    tmpHistValid   : BOOL := FALSE;
    tmpResetPrevHigh: BOOL := FALSE;
END_VAR
VAR_OUTPUT
    power      : REAL;
    correction : REAL;
    fault      : BOOL;
END_VAR
VAR_INPUT
    enable      : BOOL;
    resetBtn    : BOOL;
    sensorValid : BOOL;
    setpoint    : REAL;
    temperature : REAL;
    scanSeconds : REAL;
    bias        : REAL;
END_VAR

    (* --- Fault determination (PUB004, PUB028) --- *)
    fault := NOT sensorValid OR scanSeconds <= 0.0 OR scanSeconds > 10.0;

    (* --- Reset rising-edge detection (PUB011): edge only, not hold --- *)
    IF resetBtn AND NOT tmpResetPrevHigh THEN
        (* Rising edge of resetBtn this scan: zero outputs, clear history --- *)
        power       := 0.0;
        correction  := 0.0;
        ePrev       := 0.0;
        tmpHistValid := FALSE;
        tmpResetPrevHigh := TRUE;
        RETURN;
    END_IF

    (* Remember current resetBtn for next-scan edge detection --- *)
    tmpResetPrevHigh := resetBtn;

    (* --- Disabled or faulted: zero outputs, clear history (PUB011) --- *)
    IF NOT enable OR fault THEN
        power       := 0.0;
        correction  := 0.0;
        ePrev       := 0.0;
        tmpHistValid := FALSE;
        RETURN;
    END_IF

    (* ==================================================================
       Normal fuzzy calculation
       ================================================================== *)
    VAR
        e          : REAL;
        de         : REAL;
        x          : REAL;
        y          : REAL;
        muN_x      : REAL;
        muZ_x      : REAL;
        muP_x      : REAL;
        muN_y      : REAL;
        muZ_y      : REAL;
        muP_y      : REAL;
        w           : ARRAY[1..3, 1..3] OF REAL;
        sumW        : REAL;
        sumWc       : REAL;
        row         : INT;
        col         : INT;
        tmpFirstScan: BOOL;
    END_VAR

    (* PUB001: error definition --- *)
    e := setpoint - temperature;

    (* PUB012: first-scan detection --- *)
    tmpFirstScan := NOT tmpHistValid;

    (* PUB011: de = 0 on first scan or after history clear --- *)
    IF tmpFirstScan THEN
        de := 0.0;
    ELSE
        de := (e - ePrev) / scanSeconds;
    END_IF;

    (* PUB003 / PUB005: normalize to [-1,1] --- *)
    x := LIMIT(-1.0, e / 10.0, 1.0);
    y := LIMIT(-1.0, de / 2.0, 1.0);

    (* PUB006: membership functions --- *)
    muN_x := MAX(-x, 0.0);
    muZ_x := MAX(1.0 - ABS(x), 0.0);
    muP_x := MAX( x, 0.0);

    muN_y := MAX(-y, 0.0);
    muZ_y := MAX(1.0 - ABS(y), 0.0);
    muP_y := MAX( y, 0.0);

    (* Rule weights: row = x (N/Z/P), col = y (N/Z/P) --- *)
    w[1,1] := muN_x * muN_y;   (* N,N *)
    w[1,2] := muN_x * muZ_y;   (* N,Z *)
    w[1,3] := muN_x * muP_y;   (* N,P *)
    w[2,1] := muZ_x * muN_y;   (* Z,N *)
    w[2,2] := muZ_x * muZ_y;   (* Z,Z *)
    w[2,3] := muZ_x * muP_y;   (* Z,P *)
    w[3,1] := muP_x * muN_y;   (* P,N *)
    w[3,2] := muP_x * muZ_y;   (* P,Z *)
    w[3,3] := muP_x * muP_y;   (* P,P *)

    (* Weighted centroid (PUB007): sum(w*c)/sum(w) --- *)
    sumW  := 0.0;
    sumWc := 0.0;
    FOR row := 1 TO 3 DO
        FOR col := 1 TO 3 DO
            sumW  := sumW  + w[row, col];
            sumWc := sumWc + w[row, col] * SEL(INT_TO_INT(row - 1), SEL(INT_TO_INT(col - 1),
                                 -30.0,   (* row=1 (N) *)
                                 -10.0,   (* row=2 (Z) *)
                                  10.0),  (* row=3 (P) *)
                                 SEL(INT_TO_INT(col - 1),
                                 -20.0,   (* col=1 (N) *)
                                   0.0,   (* col=2 (Z) *)
                                  20.0)); (* col=3 (P) *)
        END_FOR;
    END_FOR;

    (* PUB007: Σw=0 → correction=0 --- *)
    IF sumW > 0.0 THEN
        correction := sumWc / sumW;
    ELSE
        correction := 0.0;
    END_IF;

    (* PUB008: power = clamp(bias + correction, 0, 100) --- *)
    power := LIMIT(0.0, bias + correction, 100.0);

    (* Update history for next scan --- *)
    ePrev       := e;
    tmpHistValid := TRUE;
END_FUNCTION_BLOCK

(* ---- self-medium-06.raw_candidate_03.st ---- *)
(* ENGINEERING_CONTRACT FB_FuzzyTempControl
   ========================================================================
   Outputs & State Retention:
   --------------------------------------------------------------------
   power:       COMBINATIONAL (bias + correction) clamped to [0,100].
                Zeroed on enable=FALSE, fault=TRUE, or resetBtn rising.
   correction:  COMBINATIONAL weighted-centroid per 9 rules.
                Zeroed same as power; no internal clamping (range ±30).
   fault:       COMBINATIONAL; fault = NOT sensorValid OR scanSeconds
                outside (0,10]. Not latched.
   ePrev:       RETAINED across scans; cleared on rising(resetBtn),
                enable=FALSE, or fault=TRUE.
   tmpHistValid:RETAINED; FALSE after clear, set TRUE after first de.
   tmpResetPrevHigh:RETAINED; set TRUE on rising(resetBtn), cleared
                next scan so held reset allows normal calculation.
   -----------------------------------------------------------------------
   First-scan rule (PUB011/PUB012): when tmpHistValid=FALSE, de=0.
   Subsequent scans use ePrev for differential calculation.
   Reset is edge-triggered only (rising edge clears; held reset allows
   normal fuzzy output per S9).
   ========================================================================
*)
FUNCTION_BLOCK FB
VAR
    ePrev          : REAL := 0.0;
    tmpHistValid   : BOOL := FALSE;
    tmpResetPrevHigh: BOOL := FALSE;
END_VAR
VAR_OUTPUT
    power      : REAL;
    correction : REAL;
    fault      : BOOL;
END_VAR
VAR_INPUT
    enable      : BOOL;
    resetBtn    : BOOL;
    sensorValid : BOOL;
    setpoint    : REAL;
    temperature : REAL;
    scanSeconds : REAL;
    bias        : REAL;
END_VAR

    (* --- Fault determination (PUB004, PUB028) --- *)
    fault := NOT sensorValid OR scanSeconds <= 0.0 OR scanSeconds > 10.0;

    (* --- Reset rising-edge detection (PUB011): edge only, not hold --- *)
    IF resetBtn AND NOT tmpResetPrevHigh THEN
        (* Rising edge of resetBtn this scan: zero outputs, clear history --- *)
        power       := 0.0;
        correction  := 0.0;
        ePrev       := 0.0;
        tmpHistValid := FALSE;
        tmpResetPrevHigh := TRUE;
        RETURN;
    END_IF;

    (* Remember current resetBtn for next-scan edge detection --- *)
    tmpResetPrevHigh := resetBtn;

    (* --- Disabled or faulted: zero outputs, clear history (PUB011) --- *)
    IF NOT enable OR fault THEN
        power       := 0.0;
        correction  := 0.0;
        ePrev       := 0.0;
        tmpHistValid := FALSE;
        RETURN;
    END_IF;

    (* ==================================================================
       Normal fuzzy calculation
       ================================================================== *)
    (* local computation variables *)
    e           : REAL;
    de          : REAL;
    x           : REAL;
    y           : REAL;
    muN_x       : REAL;
    muZ_x       : REAL;
    muP_x       : REAL;
    muN_y       : REAL;
    muZ_y       : REAL;
    muP_y       : REAL;
    w           : ARRAY[1..3, 1..3] OF REAL;
    sumW        : REAL;
    sumWc       : REAL;
    row         : INT;
    col         : INT;
    tmpFirstScan: BOOL;
END_VAR

    (* PUB001: error definition --- *)
    e := setpoint - temperature;

    (* PUB012: first-scan detection --- *)
    tmpFirstScan := NOT tmpHistValid;

    (* PUB011: de = 0 on first scan or after history clear --- *)
    IF tmpFirstScan THEN
        de := 0.0;
    ELSE
        de := (e - ePrev) / scanSeconds;
    END_IF;

    (* PUB003 / PUB005: normalize to [-1,1] --- *)
    x := LIMIT(-1.0, e / 10.0, 1.0);
    y := LIMIT(-1.0, de / 2.0, 1.0);

    (* PUB006: membership functions --- *)
    muN_x := MAX(-x, 0.0);
    muZ_x := MAX(1.0 - ABS(x), 0.0);
    muP_x := MAX( x, 0.0);

    muN_y := MAX(-y, 0.0);
    muZ_y := MAX(1.0 - ABS(y), 0.0);
    muP_y := MAX( y, 0.0);

    (* Rule weights: row = x (N/Z/P), col = y (N/Z/P) --- *)
    w[1,1] := muN_x * muN_y;   (* N,N *)
    w[1,2] := muN_x * muZ_y;   (* N,Z *)
    w[1,3] := muN_x * muP_y;   (* N,P *)
    w[2,1] := muZ_x * muN_y;   (* Z,N *)
    w[2,2] := muZ_x * muZ_y;   (* Z,Z *)
    w[2,3] := muZ_x * muP_y;   (* Z,P *)
    w[3,1] := muP_x * muN_y;   (* P,N *)
    w[3,2] := muP_x * muZ_y;   (* P,Z *)
    w[3,3] := muP_x * muP_y;   (* P,P *)

    (* Weighted centroid (PUB007): sum(w*c)/sum(w) --- *)
    sumW  := 0.0;
    sumWc := 0.0;
    FOR row := 1 TO 3 DO
        FOR col := 1 TO 3 DO
            sumW  := sumW  + w[row, col];
            sumWc := sumWc + w[row, col] * SEL(INT_TO_INT(row - 1), SEL(INT_TO_INT(col - 1),
                                 -30.0,   (* row=1 (N) *)
                                 -10.0,   (* row=2 (Z) *)
                                  10.0),  (* row=3 (P) *)
                                 SEL(INT_TO_INT(col - 1),
                                 -20.0,   (* col=1 (N) *)
                                   0.0,   (* col=2 (Z) *)
                                  20.0)); (* col=3 (P) *)
        END_FOR;
    END_FOR;

    (* PUB007: Σw=0 → correction=0 --- *)
    IF sumW > 0.0 THEN
        correction := sumWc / sumW;
    ELSE
        correction := 0.0;
    END_IF;

    (* PUB008: power = clamp(bias + correction, 0, 100) --- *)
    power := LIMIT(0.0, bias + correction, 100.0);

    (* Update history for next scan --- *)
    ePrev       := e;
    tmpHistValid := TRUE;
END_FUNCTION_BLOCK

(* ---- self-medium-06.raw_candidate_04.st ---- *)
(* ENGINEERING_CONTRACT FB_FuzzyTempControl
   ========================================================================
   Outputs & State Retention:
   --------------------------------------------------------------------
   power:       COMBINATIONAL (bias + correction) clamped to [0,100].
                Zeroed on enable=FALSE, fault=TRUE, or resetBtn rising.
   correction:  COMBINATIONAL weighted-centroid per 9 rules.
                Zeroed same as power; no internal clamping (range ±30).
   fault:       COMBINATIONAL; fault = NOT sensorValid OR scanSeconds
                outside (0,10]. Not latched.
   ePrev:       RETAINED across scans; cleared on rising(resetBtn),
                enable=FALSE, or fault=TRUE.
   tmpHistValid:RETAINED; FALSE after clear, set TRUE after first de.
   tmpResetPrevHigh:RETAINED; set TRUE on rising(resetBtn), cleared
                next scan so held reset allows normal calculation.
   -----------------------------------------------------------------------
   First-scan rule (PUB011/PUB012): when tmpHistValid=FALSE, de=0.
   Subsequent scans use ePrev for differential calculation.
   Reset is edge-triggered only (rising edge clears; held reset allows
   normal fuzzy output per S9).
   ========================================================================
*)
FUNCTION_BLOCK FB
VAR
    ePrev           : REAL := 0.0;
    tmpHistValid    : BOOL := FALSE;
    tmpResetPrevHigh: BOOL := FALSE;
    e               : REAL;
    de              : REAL;
    x               : REAL;
    y               : REAL;
    muN_x           : REAL;
    muZ_x           : REAL;
    muP_x           : REAL;
    muN_y           : REAL;
    muZ_y           : REAL;
    muP_y           : REAL;
    w               : ARRAY[1..3, 1..3] OF REAL;
    sumW            : REAL;
    sumWc           : REAL;
    row             : INT;
    col             : INT;
    tmpFirstScan    : BOOL;
END_VAR
VAR_OUTPUT
    power      : REAL;
    correction : REAL;
    fault      : BOOL;
END_VAR
VAR_INPUT
    enable      : BOOL;
    resetBtn    : BOOL;
    sensorValid : BOOL;
    setpoint    : REAL;
    temperature : REAL;
    scanSeconds : REAL;
    bias        : REAL;
END_VAR

    (* --- Fault determination (PUB004, PUB028) --- *)
    fault := NOT sensorValid OR scanSeconds <= 0.0 OR scanSeconds > 10.0;

    (* --- Reset rising-edge detection (PUB011): edge only, not hold --- *)
    IF resetBtn AND NOT tmpResetPrevHigh THEN
        (* Rising edge of resetBtn this scan: zero outputs, clear history --- *)
        power        := 0.0;
        correction   := 0.0;
        ePrev        := 0.0;
        tmpHistValid := FALSE;
        tmpResetPrevHigh := TRUE;
        RETURN;
    END_IF;

    (* Remember current resetBtn for next-scan edge detection --- *)
    tmpResetPrevHigh := resetBtn;

    (* --- Disabled or faulted: zero outputs, clear history (PUB011) --- *)
    IF NOT enable OR fault THEN
        power        := 0.0;
        correction   := 0.0;
        ePrev        := 0.0;
        tmpHistValid := FALSE;
        RETURN;
    END_IF;

    (* ==================================================================
       Normal fuzzy calculation
       ================================================================== *)

    (* PUB001: error definition --- *)
    e := setpoint - temperature;

    (* PUB012: first-scan detection --- *)
    tmpFirstScan := NOT tmpHistValid;

    (* PUB011: de = 0 on first scan or after history clear --- *)
    IF tmpFirstScan THEN
        de := 0.0;
    ELSE
        de := (e - ePrev) / scanSeconds;
    END_IF;

    (* PUB003 / PUB005: normalize to [-1,1] --- *)
    x := LIMIT(-1.0, e / 10.0, 1.0);
    y := LIMIT(-1.0, de / 2.0, 1.0);

    (* PUB006: membership functions --- *)
    muN_x := MAX(-x, 0.0);
    muZ_x := MAX(1.0 - ABS(x), 0.0);
    muP_x := MAX( x, 0.0);

    muN_y := MAX(-y, 0.0);
    muZ_y := MAX(1.0 - ABS(y), 0.0);
    muP_y := MAX( y, 0.0);

    (* Rule weights: row = x (N/Z/P), col = y (N/Z/P) --- *)
    w[1,1] := muN_x * muN_y;   (* N,N *)
    w[1,2] := muN_x * muZ_y;   (* N,Z *)
    w[1,3] := muN_x * muP_y;   (* N,P *)
    w[2,1] := muZ_x * muN_y;   (* Z,N *)
    w[2,2] := muZ_x * muZ_y;   (* Z,Z *)
    w[2,3] := muZ_x * muP_y;   (* Z,P *)
    w[3,1] := muP_x * muN_y;   (* P,N *)
    w[3,2] := muP_x * muZ_y;   (* P,Z *)
    w[3,3] := muP_x * muP_y;   (* P,P *)

    (* Weighted centroid (PUB007): sum(w*c)/sum(w) --- *)
    sumW  := 0.0;
    sumWc := 0.0;
    FOR row := 1 TO 3 DO
        FOR col := 1 TO 3 DO
            sumW  := sumW  + w[row, col];
            sumWc := sumWc + w[row, col] * SEL(INT_TO_INT(row - 1), SEL(INT_TO_INT(col - 1),
                                 -30.0,   (* row=1 (N) *)
                                 -10.0,   (* row=2 (Z) *)
                                  10.0),  (* row=3 (P) *)
                                 SEL(INT_TO_INT(col - 1),
                                 -20.0,   (* col=1 (N) *)
                                   0.0,   (* col=2 (Z) *)
                                  20.0)); (* col=3 (P) *)
        END_FOR;
    END_FOR;

    (* PUB007: Σw=0 → correction=0 --- *)
    IF sumW > 0.0 THEN
        correction := sumWc / sumW;
    ELSE
        correction := 0.0;
    END_IF;

    (* PUB008: power = clamp(bias + correction, 0, 100) --- *)
    power := LIMIT(0.0, bias + correction, 100.0);

    (* Update history for next scan --- *)
    ePrev        := e;
    tmpHistValid := TRUE;
END_FUNCTION_BLOCK
